(* IEC 61131-3 sources: kns-pump-station/tests/POUs/Model/FB_VfdSim_Test, 29 files *)

(* ---- FB_VfdSim_Test.decl.st ---- *)
// Назначение: набор coUnit для FB_VfdSim — модель ПЧ по условной карте: рампа к заданию и торможение, реле
//             «Работа», авария с выбегом и сброс по фронту CTW.2, коды аварий, потеря связи (регистры замирают,
//             записи не доходят), сторожевой таймер 5 с → 50 Гц (04 §12, PMI-28, PMI-29), восстановление связи,
//             пропадание питания и загрузка, инъекции ОС, местный пуск (частота местного поста), ток в регистре,
//             «время назад».
//             Время — PL.FB_FakeTime, шаг 100 мс; разгон 0 → 50 Гц за 10 с (5 Гц/с).
// Автор:      kr0nsch
// Версия:     0.1.0
// Документ:   docs/DESIGN.md, разделы 11.3, 14.1
FUNCTION_BLOCK FB_VfdSim_Test EXTENDS coUnit.FB_TestSuite
VAR CONSTANT
    T_STEP : TIME := T#100MS;
    UI_1S : UINT := 10;               // шагов в 1 с
    R_EPS_HZ : REAL := 1.0E-3;
    UI_FREF_50HZ : UINT := 5000;      // 0,01 Гц
    UI_FREF_30HZ : UINT := 3000;
    UI_FREF_25HZ : UINT := 2500;
    R_LOCAL_HZ : REAL := 50.0;        // частота местного поста (SIM_VFD_LOCAL_FREQ_HZ)
END_VAR

(* ---- CommLossFreezesRegisters.method.decl.st ---- *)
// Потеря связи на 25 Гц: xCommOk = FALSE, регистры STW и FACT замирают; новое задание не доходит
// (частота 25 Гц); стоп по проводу работает (через 2 с — 15 Гц), а FACT по-прежнему 2500.
METHOD PRIVATE CommLossFreezesRegisters
VAR
    fbTime : PL.FB_FakeTime;    // подменное время
    fbDut : FB_VfdSim;          // проверяемая модель ПЧ
    uiI : UINT;
END_VAR

(* ---- CommLossFreezesRegisters.method.impl.st ---- *)
coUnit.TEST('VfdSim_CommLossFreezesRegisters');

fbDut(xRunCmd := TRUE, uiFref := UI_FREF_25HZ, itfTime := fbTime);
FOR uiI := 1 TO 6 * UI_1S DO
    fbTime.Advance(tStep := T_STEP);
    fbDut(itfTime := fbTime);
END_FOR
AssertEquals_UINT(Expected := 2500, Actual := fbDut.uiFact, Message := 'FACT 2500 before loss');
fbDut.xCommLoss := TRUE;
FOR uiI := 1 TO 1 DO
    fbTime.Advance(tStep := T_STEP);
    fbDut(itfTime := fbTime);
END_FOR
AssertFalse(Condition := fbDut.xCommOk, Message := 'no comm');
fbDut.uiFref := UI_FREF_50HZ;
FOR uiI := 1 TO 2 * UI_1S DO
    fbTime.Advance(tStep := T_STEP);
    fbDut(itfTime := fbTime);
END_FOR
AssertEquals_REAL(Expected := 25.0, Actual := fbDut.rFreq_Hz, Delta := R_EPS_HZ,
                  Message := 'new reference not received');
fbDut.xRunCmd := FALSE;
FOR uiI := 1 TO 2 * UI_1S DO
    fbTime.Advance(tStep := T_STEP);
    fbDut(itfTime := fbTime);
END_FOR
AssertEquals_REAL(Expected := 15.0, Actual := fbDut.rFreq_Hz, Delta := R_EPS_HZ, Message := 'wired stop works');
AssertEquals_UINT(Expected := 2500, Actual := fbDut.uiFact, Message := 'FACT frozen');
AssertEquals_WORD(Expected := GVL_Const.VFD_STW_READY OR GVL_Const.VFD_STW_RUNNING OR GVL_Const.VFD_STW_REMOTE,
                  Actual := fbDut.wStw, Message := 'STW frozen');

coUnit.TEST_FINISHED();

(* ---- CommLossWatchdogGoesTo50HzAfter5s.method.decl.st ---- *)
// Сторожевой таймер ПЧ (04 §12): работающий на 30 Гц насос через 4,9 с без связи — ещё задание 30 Гц,
// в 5,0 с — 50 Гц, через 4 с разгона — 50 Гц. Стоящий насос без связи (последнее задание 0): пуск по
// проводу после срабатывания таймера — разгон до 50 Гц, а не работа на 0 Гц.
METHOD PRIVATE CommLossWatchdogGoesTo50HzAfter5s
VAR
    fbTime : PL.FB_FakeTime;    // подменное время
    fbDut : FB_VfdSim;          // проверяемая модель ПЧ
    uiI : UINT;
    fbStopped : FB_VfdSim;      // ПЧ стоящего насоса
END_VAR

(* ---- CommLossWatchdogGoesTo50HzAfter5s.method.impl.st ---- *)
coUnit.TEST('VfdSim_CommLossWatchdogGoesTo50HzAfter5s');

fbDut(xRunCmd := TRUE, uiFref := UI_FREF_30HZ, itfTime := fbTime);
fbStopped(xRunCmd := FALSE, uiFref := 0, itfTime := fbTime);
FOR uiI := 1 TO 6 * UI_1S DO
    fbTime.Advance(tStep := T_STEP);
    fbDut(itfTime := fbTime);
END_FOR
fbDut.xCommLoss := TRUE;
fbStopped.xCommLoss := TRUE;
fbTime.Advance(tStep := T_STEP);
fbDut(itfTime := fbTime);
fbStopped(itfTime := fbTime);
FOR uiI := 1 TO 5 * UI_1S - 1 DO
    fbTime.Advance(tStep := T_STEP);
    fbDut(itfTime := fbTime);
    fbStopped(itfTime := fbTime);
END_FOR
AssertFalse(Condition := fbDut.xWatchdog, Message := 'no watchdog at 4.9 s');
AssertEquals_REAL(Expected := 30.0, Actual := fbDut.rRef_Hz, Delta := R_EPS_HZ, Message := 'last reference 30 Hz');
fbTime.Advance(tStep := T_STEP);
fbDut(itfTime := fbTime);
fbStopped(itfTime := fbTime);
AssertTrue(Condition := fbDut.xWatchdog AND fbStopped.xWatchdog, Message := 'watchdog at 5.0 s');
AssertEquals_REAL(Expected := GVL_Const.SIM_VFD_WATCHDOG_FREQ_HZ, Actual := fbDut.rRef_Hz, Delta := 0.0,
                  Message := 'preset 50 Hz');
FOR uiI := 1 TO 10 * UI_1S DO
    fbTime.Advance(tStep := T_STEP);
    fbDut(itfTime := fbTime);
    fbStopped(xRunCmd := TRUE, itfTime := fbTime);
END_FOR
AssertEquals_REAL(Expected := 50.0, Actual := fbDut.rFreq_Hz, Delta := R_EPS_HZ, Message := 'running pump at 50 Hz');
AssertEquals_REAL(Expected := 50.0, Actual := fbStopped.rFreq_Hz, Delta := R_EPS_HZ,
                  Message := 'pump started by wire runs at 50 Hz');

coUnit.TEST_FINISHED();

(* ---- CommRestoredFollowsFref.method.decl.st ---- *)
// После срабатывания таймера (50 Гц) связь восстановлена с заданием 3000: таймер снят, задание 30 Гц,
// через 4 с — 30 Гц, регистры снова обновляются (FACT 3000).
METHOD PRIVATE CommRestoredFollowsFref
VAR
    fbTime : PL.FB_FakeTime;    // подменное время
    fbDut : FB_VfdSim;          // проверяемая модель ПЧ
    uiI : UINT;
END_VAR

(* ---- CommRestoredFollowsFref.method.impl.st ---- *)
coUnit.TEST('VfdSim_CommRestoredFollowsFref');

fbDut(xRunCmd := TRUE, uiFref := UI_FREF_50HZ, itfTime := fbTime);
FOR uiI := 1 TO 10 * UI_1S DO
    fbTime.Advance(tStep := T_STEP);
    fbDut(itfTime := fbTime);
END_FOR
fbDut.xCommLoss := TRUE;
FOR uiI := 1 TO 6 * UI_1S DO
    fbTime.Advance(tStep := T_STEP);
    fbDut(itfTime := fbTime);
END_FOR
AssertTrue(Condition := fbDut.xWatchdog, Message := 'watchdog active');
fbDut.xCommLoss := FALSE;
fbDut.uiFref := UI_FREF_30HZ;
FOR uiI := 1 TO 1 DO
    fbTime.Advance(tStep := T_STEP);
    fbDut(itfTime := fbTime);
END_FOR
AssertTrue(Condition := fbDut.xCommOk AND NOT fbDut.xWatchdog, Message := 'comm restored, watchdog off');
AssertEquals_REAL(Expected := 30.0, Actual := fbDut.rRef_Hz, Delta := R_EPS_HZ, Message := 'follows FREF again');
FOR uiI := 1 TO 4 * UI_1S DO
    fbTime.Advance(tStep := T_STEP);
    fbDut(itfTime := fbTime);
END_FOR
AssertEquals_REAL(Expected := 30.0, Actual := fbDut.rFreq_Hz, Delta := R_EPS_HZ, Message := 'ramped to 30 Hz');
AssertEquals_UINT(Expected := 3000, Actual := fbDut.uiFact, Message := 'FACT updated');

coUnit.TEST_FINISHED();

(* ---- CurrentRegisterScaled.method.decl.st ---- *)
// Ток двигателя в регистре 102 — 0,1 А: 26,38 А → 264; неконечный ток и стоящий ПЧ — 0.
METHOD PRIVATE CurrentRegisterScaled
VAR
    fbTime : PL.FB_FakeTime;    // подменное время
    fbDut : FB_VfdSim;          // проверяемая модель ПЧ
    uiI : UINT;
    uBits : PL.U_RealBits;
END_VAR

(* ---- CurrentRegisterScaled.method.impl.st ---- *)
coUnit.TEST('VfdSim_CurrentRegisterScaled');

fbDut(xRunCmd := TRUE, uiFref := UI_FREF_50HZ, itfTime := fbTime);
FOR uiI := 1 TO 10 * UI_1S DO
    fbTime.Advance(tStep := T_STEP);
    fbDut(itfTime := fbTime);
END_FOR
fbDut.rMotorCurrent_A := 26.38;
FOR uiI := 1 TO 1 DO
    fbTime.Advance(tStep := T_STEP);
    fbDut(itfTime := fbTime);
END_FOR
AssertEquals_UINT(Expected := 264, Actual := fbDut.uiCurrent, Message := '26.38 A -> 264');
uBits.dwValue := 16#7FC00000;
fbDut.rMotorCurrent_A := uBits.rValue;
FOR uiI := 1 TO 1 DO
    fbTime.Advance(tStep := T_STEP);
    fbDut(itfTime := fbTime);
END_FOR
AssertEquals_UINT(Expected := 0, Actual := fbDut.uiCurrent, Message := 'NaN current -> 0');
fbDut.rMotorCurrent_A := 26.38;
fbDut.xRunCmd := FALSE;
FOR uiI := 1 TO 11 * UI_1S DO
    fbTime.Advance(tStep := T_STEP);
    fbDut(itfTime := fbTime);
END_FOR
AssertEquals_UINT(Expected := 0, Actual := fbDut.uiCurrent, Message := 'stopped drive -> 0');

coUnit.TEST_FINISHED();

(* ---- DefaultsReadyAndStopped.method.decl.st ---- *)
// Первый вызов с питанием: ПЧ готов, связь есть, STW = готов + дистанционное (16#0011), частота и
// FACT 0, код аварии 0, реле разомкнуты.
METHOD PRIVATE DefaultsReadyAndStopped
VAR
    fbTime : PL.FB_FakeTime;    // подменное время
    fbDut : FB_VfdSim;          // проверяемая модель ПЧ
END_VAR

(* ---- FaultCoastAndResetEdge.method.decl.st ---- *)
// Авария ПЧ на 50 Гц: выбег (частота 0 сразу), реле «Авария», STW.2, код 11, не готов. Сброс при
// активной инъекции не снимает; после снятия инъекции нужен новый фронт CTW.2; код аварии остаётся.
METHOD PRIVATE FaultCoastAndResetEdge
VAR
    fbTime : PL.FB_FakeTime;    // подменное время
    fbDut : FB_VfdSim;          // проверяемая модель ПЧ
    uiI : UINT;
END_VAR

(* ---- FaultCoastAndResetEdge.method.impl.st ---- *)
coUnit.TEST('VfdSim_FaultCoastAndResetEdge');

fbDut(xRunCmd := TRUE, uiFref := UI_FREF_50HZ, itfTime := fbTime);
FOR uiI := 1 TO 10 * UI_1S DO
    fbTime.Advance(tStep := T_STEP);
    fbDut(itfTime := fbTime);
END_FOR
fbDut.xFaultInj := TRUE;
FOR uiI := 1 TO 1 DO
    fbTime.Advance(tStep := T_STEP);
    fbDut(itfTime := fbTime);
END_FOR
AssertEquals_REAL(Expected := 0.0, Actual := fbDut.rFreq_Hz, Delta := 0.0, Message := 'coast: frequency 0');
AssertTrue(Condition := fbDut.xRelayFault AND fbDut.xFaulted AND NOT fbDut.xReady, Message := 'fault latched');
AssertFalse(Condition := fbDut.xRelayRun, Message := 'run relay open');
AssertEquals_WORD(Expected := GVL_Const.VFD_STW_FAULT OR GVL_Const.VFD_STW_REMOTE, Actual := fbDut.wStw,
                  Message := 'STW fault + remote');
AssertEquals_UINT(Expected := GVL_Const.SIM_VFD_FCODE_EXT, Actual := fbDut.uiFcode, Message := 'fault code 11');
fbDut.wCtw := GVL_Const.VFD_CTW_RESET;
FOR uiI := 1 TO 1 DO
    fbTime.Advance(tStep := T_STEP);
    fbDut(itfTime := fbTime);
END_FOR
AssertTrue(Condition := fbDut.xFaulted, Message := 'reset ignored while cause active');
fbDut.xFaultInj := FALSE;
FOR uiI := 1 TO 1 DO
    fbTime.Advance(tStep := T_STEP);
    fbDut(itfTime := fbTime);
END_FOR
AssertTrue(Condition := fbDut.xFaulted, Message := 'no new reset edge: still faulted');
fbDut.wCtw := 0;
FOR uiI := 1 TO 1 DO
    fbTime.Advance(tStep := T_STEP);
    fbDut(itfTime := fbTime);
END_FOR
fbDut.wCtw := GVL_Const.VFD_CTW_RESET;
FOR uiI := 1 TO 1 DO
    fbTime.Advance(tStep := T_STEP);
    fbDut(itfTime := fbTime);
END_FOR
AssertFalse(Condition := fbDut.xFaulted OR fbDut.xRelayFault, Message := 'reset edge clears fault');
AssertTrue(Condition := fbDut.xReady, Message := 'ready again');
AssertEquals_UINT(Expected := GVL_Const.SIM_VFD_FCODE_EXT, Actual := fbDut.uiFcode, Message := 'last fault code kept');
FOR uiI := 1 TO 1 DO
    fbTime.Advance(tStep := T_STEP);
    fbDut(itfTime := fbTime);
END_FOR
AssertTrue(Condition := fbDut.xOutputActive AND fbDut.rFreq_Hz > 0.0, Message := 'wired run restarts the drive');

coUnit.TEST_FINISHED();

(* ---- FeedbackStuckInjection.method.decl.st ---- *)
// Инъекция «ОС залипла»: ПЧ стоит, реле «Работа» замкнуто.
METHOD PRIVATE FeedbackStuckInjection
VAR
    fbTime : PL.FB_FakeTime;    // подменное время
    fbDut : FB_VfdSim;          // проверяемая модель ПЧ
END_VAR

(* ---- LocalRun.method.decl.st ---- *)
// «Местное»: провод «Пуск» от ПЛК не действует, пуск — с местного поста; бит STW.4 (дистанционное)
// снят.
METHOD PRIVATE LocalRun
VAR
    fbTime : PL.FB_FakeTime;    // подменное время
    fbDut : FB_VfdSim;          // проверяемая модель ПЧ
    uiI : UINT;
END_VAR

(* ---- LocalRun.method.impl.st ---- *)
coUnit.TEST('VfdSim_LocalRun');

fbDut(xRunCmd := TRUE, xLocal := TRUE, uiFref := UI_FREF_50HZ, itfTime := fbTime);
FOR uiI := 1 TO UI_1S DO
    fbTime.Advance(tStep := T_STEP);
    fbDut(itfTime := fbTime);
END_FOR
AssertFalse(Condition := fbDut.xOutputActive, Message := 'PLC wire ignored in local');
AssertEquals_WORD(Expected := GVL_Const.VFD_STW_READY, Actual := fbDut.wStw, Message := 'STW without remote bit');
fbDut.xLocalRun := TRUE;
FOR uiI := 1 TO UI_1S DO
    fbTime.Advance(tStep := T_STEP);
    fbDut(itfTime := fbTime);
END_FOR
AssertTrue(Condition := fbDut.xOutputActive AND fbDut.xRelayRun, Message := 'local run starts the drive');
AssertEquals_REAL(Expected := 5.0, Actual := fbDut.rFreq_Hz, Delta := R_EPS_HZ, Message := 'ramp in local');

coUnit.TEST_FINISHED();

(* ---- LocalRunAtLocalPreset.method.decl.st ---- *)
// «Местное», пуск по месту у стоящего насоса: FB_MotorVfd в Local держит задание равным фактической
// скорости (0 % у стоящего насоса), FREF = 0. ПЧ разгоняется к частоте местного поста (50 Гц) за tAccel,
// записи FREF мастера в «Местном» не действуют; после возврата в «Дистанционное» — снова FREF.
METHOD PRIVATE LocalRunAtLocalPreset
VAR
    fbTime : PL.FB_FakeTime;    // подменное время
    fbDut : FB_VfdSim;          // проверяемая модель ПЧ
    uiI : UINT;
END_VAR

(* ---- LocalRunAtLocalPreset.method.impl.st ---- *)
coUnit.TEST('VfdSim_LocalRunAtLocalPreset');

fbDut(xLocal := TRUE, xLocalRun := TRUE, uiFref := 0, itfTime := fbTime);
FOR uiI := 1 TO 10 * UI_1S DO
    fbTime.Advance(tStep := T_STEP);
    fbDut(itfTime := fbTime);
END_FOR
AssertTrue(Condition := fbDut.xOutputActive AND fbDut.xRelayRun, Message := 'local run starts the drive');
AssertEquals_REAL(Expected := R_LOCAL_HZ, Actual := fbDut.rFreq_Hz, Delta := R_EPS_HZ,
                  Message := 'local preset reached in tAccel');
fbDut.uiFref := UI_FREF_25HZ;
FOR uiI := 1 TO UI_1S DO
    fbTime.Advance(tStep := T_STEP);
    fbDut(itfTime := fbTime);
END_FOR
AssertEquals_REAL(Expected := R_LOCAL_HZ, Actual := fbDut.rFreq_Hz, Delta := R_EPS_HZ,
                  Message := 'master FREF ignored in local');
fbDut.xLocal := FALSE;
fbDut.xLocalRun := FALSE;
fbDut.xRunCmd := TRUE;
FOR uiI := 1 TO 5 * UI_1S DO
    fbTime.Advance(tStep := T_STEP);
    fbDut(itfTime := fbTime);
END_FOR
AssertEquals_REAL(Expected := 25.0, Actual := fbDut.rFreq_Hz, Delta := R_EPS_HZ, Message := 'remote: back to FREF');

coUnit.TEST_FINISHED();

(* ---- NoFeedbackInjection.method.decl.st ---- *)
// Инъекция «нет ОС»: ПЧ вращает насос, реле «Работа» разомкнуто.
METHOD PRIVATE NoFeedbackInjection
VAR
    fbTime : PL.FB_FakeTime;    // подменное время
    fbDut : FB_VfdSim;          // проверяемая модель ПЧ
    uiI : UINT;
END_VAR

(* ---- NoFeedbackInjection.method.impl.st ---- *)
coUnit.TEST('VfdSim_NoFeedbackInjection');

fbDut(xRunCmd := TRUE, uiFref := UI_FREF_50HZ, itfTime := fbTime);
FOR uiI := 1 TO 10 * UI_1S DO
    fbTime.Advance(tStep := T_STEP);
    fbDut(itfTime := fbTime);
END_FOR
fbDut.xNoFeedback := TRUE;
FOR uiI := 1 TO 1 DO
    fbTime.Advance(tStep := T_STEP);
    fbDut(itfTime := fbTime);
END_FOR
AssertTrue(Condition := fbDut.rFreq_Hz > 0.0 AND fbDut.xOutputActive, Message := 'drive running');
AssertFalse(Condition := fbDut.xRelayRun, Message := 'run relay open (no feedback)');

coUnit.TEST_FINISHED();

(* ---- OverheatFaultCode.method.decl.st ---- *)
// Перегрев (TS1n2 разрывает цепь аварии): авария ПЧ с кодом 12, выбег.
METHOD PRIVATE OverheatFaultCode
VAR
    fbTime : PL.FB_FakeTime;    // подменное время
    fbDut : FB_VfdSim;          // проверяемая модель ПЧ
    uiI : UINT;
END_VAR

(* ---- OverheatFaultCode.method.impl.st ---- *)
coUnit.TEST('VfdSim_OverheatFaultCode');

fbDut(xRunCmd := TRUE, uiFref := UI_FREF_50HZ, itfTime := fbTime);
FOR uiI := 1 TO 10 * UI_1S DO
    fbTime.Advance(tStep := T_STEP);
    fbDut(itfTime := fbTime);
END_FOR
fbDut.xOverheat := TRUE;
FOR uiI := 1 TO 1 DO
    fbTime.Advance(tStep := T_STEP);
    fbDut(itfTime := fbTime);
END_FOR
AssertTrue(Condition := fbDut.xFaulted AND fbDut.xRelayFault, Message := 'overheat trips the drive');
AssertEquals_UINT(Expected := GVL_Const.SIM_VFD_FCODE_OVERHEAT, Actual := fbDut.uiFcode, Message := 'fault code 12');
AssertEquals_REAL(Expected := 0.0, Actual := fbDut.rFreq_Hz, Delta := 0.0, Message := 'coast');

coUnit.TEST_FINISHED();

(* ---- PowerLossAndBoot.method.decl.st ---- *)
// Пропадание питания на ходу: частота 0, реле разомкнуты, связи нет, регистры 0. Питание вернулось
// (первый шаг цикла — вызов с питанием): 4,9 с ПЧ загружается (STW 0, связи нет), в 5,0 с готов, код
// последней аварии 13 (пониженное напряжение), пуск по проводу удержан — разгон.
METHOD PRIVATE PowerLossAndBoot
VAR
    fbTime : PL.FB_FakeTime;    // подменное время
    fbDut : FB_VfdSim;          // проверяемая модель ПЧ
    uiI : UINT;
END_VAR

(* ---- PowerLossAndBoot.method.impl.st ---- *)
coUnit.TEST('VfdSim_PowerLossAndBoot');

fbDut(xRunCmd := TRUE, uiFref := UI_FREF_50HZ, itfTime := fbTime);
FOR uiI := 1 TO 10 * UI_1S DO
    fbTime.Advance(tStep := T_STEP);
    fbDut(itfTime := fbTime);
END_FOR
fbDut.xPowerOk := FALSE;
FOR uiI := 1 TO 1 DO
    fbTime.Advance(tStep := T_STEP);
    fbDut(itfTime := fbTime);
END_FOR
AssertEquals_REAL(Expected := 0.0, Actual := fbDut.rFreq_Hz, Delta := 0.0, Message := 'no power: frequency 0');
AssertFalse(Condition := fbDut.xRelayRun OR fbDut.xCommOk OR fbDut.xReady, Message := 'no power: relays, comm off');
AssertEquals_WORD(Expected := 0, Actual := fbDut.wStw, Message := 'no power: STW 0');
fbDut.xPowerOk := TRUE;
FOR uiI := 1 TO 5 * UI_1S DO
    fbTime.Advance(tStep := T_STEP);
    fbDut(itfTime := fbTime);
END_FOR
AssertFalse(Condition := fbDut.xReady OR fbDut.xCommOk, Message := 'booting at 4.9 s');
AssertEquals_WORD(Expected := 0, Actual := fbDut.wStw, Message := 'booting: STW 0');
FOR uiI := 1 TO 1 DO
    fbTime.Advance(tStep := T_STEP);
    fbDut(itfTime := fbTime);
END_FOR
AssertTrue(Condition := fbDut.xReady AND fbDut.xCommOk, Message := 'ready after boot');
AssertEquals_UINT(Expected := GVL_Const.SIM_VFD_FCODE_UNDERVOLT, Actual := fbDut.uiFcode,
                  Message := 'last fault: undervoltage');
AssertTrue(Condition := fbDut.xOutputActive, Message := 'held wired run restarts after boot');

coUnit.TEST_FINISHED();

(* ---- RampToReference.method.decl.st ---- *)
// Пуск с заданием 5000 (50 Гц): через 5 с — 25 Гц (FACT 2500), через 10 с — 50 Гц; реле «Работа»
// и бит STW.1. Стоп: торможение 5 Гц/с, реле замкнуто до остановки (через 9,9 с — 0,5 Гц), в 10 с — 0.
METHOD PRIVATE RampToReference
VAR
    fbTime : PL.FB_FakeTime;    // подменное время
    fbDut : FB_VfdSim;          // проверяемая модель ПЧ
    uiI : UINT;
END_VAR

(* ---- RampToReference.method.impl.st ---- *)
coUnit.TEST('VfdSim_RampToReference');

fbDut(xRunCmd := TRUE, uiFref := UI_FREF_50HZ, itfTime := fbTime);
FOR uiI := 1 TO 5 * UI_1S DO
    fbTime.Advance(tStep := T_STEP);
    fbDut(itfTime := fbTime);
END_FOR
AssertEquals_REAL(Expected := 25.0, Actual := fbDut.rFreq_Hz, Delta := R_EPS_HZ, Message := '25 Hz after 5 s');
AssertEquals_UINT(Expected := 2500, Actual := fbDut.uiFact, Message := 'FACT 2500');
AssertTrue(Condition := fbDut.xRelayRun, Message := 'run relay closed');
AssertEquals_WORD(Expected := GVL_Const.VFD_STW_READY OR GVL_Const.VFD_STW_RUNNING OR GVL_Const.VFD_STW_REMOTE,
                  Actual := fbDut.wStw, Message := 'STW ready + running + remote');
FOR uiI := 1 TO 5 * UI_1S DO
    fbTime.Advance(tStep := T_STEP);
    fbDut(itfTime := fbTime);
END_FOR
AssertEquals_REAL(Expected := 50.0, Actual := fbDut.rFreq_Hz, Delta := R_EPS_HZ, Message := '50 Hz after 10 s');
AssertEquals_UINT(Expected := 5000, Actual := fbDut.uiFact, Message := 'FACT 5000');
fbDut.xRunCmd := FALSE;
FOR uiI := 1 TO 10 * UI_1S - 1 DO
    fbTime.Advance(tStep := T_STEP);
    fbDut(itfTime := fbTime);
END_FOR
AssertEquals_REAL(Expected := 0.5, Actual := fbDut.rFreq_Hz, Delta := R_EPS_HZ, Message := 'decelerating: 0.5 Hz');
AssertTrue(Condition := fbDut.xRelayRun, Message := 'run relay closed while decelerating');
FOR uiI := 1 TO 1 DO
    fbTime.Advance(tStep := T_STEP);
    fbDut(itfTime := fbTime);
END_FOR
AssertEquals_REAL(Expected := 0.0, Actual := fbDut.rFreq_Hz, Delta := 0.0, Message := 'stopped');
AssertFalse(Condition := fbDut.xRelayRun OR fbDut.xOutputActive, Message := 'run relay open after stop');

coUnit.TEST_FINISHED();

(* ---- ResetDriveClearsFault.method.decl.st ---- *)
// ResetDrive («ПЧ готовы», xResetPlant) снимает аварию, если причины уже нет, без фронта CTW.2;
// при активной причине авария остаётся.
METHOD PRIVATE ResetDriveClearsFault
VAR
    fbTime : PL.FB_FakeTime;    // подменное время
    fbDut : FB_VfdSim;          // проверяемая модель ПЧ
    uiI : UINT;
END_VAR

(* ---- ResetDriveClearsFault.method.impl.st ---- *)
coUnit.TEST('VfdSim_ResetDriveClearsFault');

fbDut(xRunCmd := TRUE, uiFref := UI_FREF_50HZ, itfTime := fbTime);
FOR uiI := 1 TO 10 * UI_1S DO
    fbTime.Advance(tStep := T_STEP);
    fbDut(itfTime := fbTime);
END_FOR
fbDut.xFaultInj := TRUE;
FOR uiI := 1 TO 1 DO
    fbTime.Advance(tStep := T_STEP);
    fbDut(itfTime := fbTime);
END_FOR
fbDut.ResetDrive();
FOR uiI := 1 TO 1 DO
    fbTime.Advance(tStep := T_STEP);
    fbDut(itfTime := fbTime);
END_FOR
AssertTrue(Condition := fbDut.xFaulted, Message := 'cause active: fault stays');
fbDut.xFaultInj := FALSE;
fbDut.ResetDrive();
FOR uiI := 1 TO 1 DO
    fbTime.Advance(tStep := T_STEP);
    fbDut(itfTime := fbTime);
END_FOR
AssertFalse(Condition := fbDut.xFaulted, Message := 'ResetDrive clears fault');
AssertTrue(Condition := fbDut.xReady, Message := 'ready');

coUnit.TEST_FINISHED();

(* ---- TimeBackwardsHoldsFrequency.method.decl.st ---- *)
// «Время назад»: шаг рампы 0 — частота не меняется; дальше рампа продолжается.
METHOD PRIVATE TimeBackwardsHoldsFrequency
VAR
    fbTime : PL.FB_FakeTime;    // подменное время
    fbDut : FB_VfdSim;          // проверяемая модель ПЧ
    uiI : UINT;
END_VAR

(* ---- TimeBackwardsHoldsFrequency.method.impl.st ---- *)
coUnit.TEST('VfdSim_TimeBackwardsHoldsFrequency');

fbDut(xRunCmd := TRUE, uiFref := UI_FREF_50HZ, itfTime := fbTime);
FOR uiI := 1 TO 3 * UI_1S DO
    fbTime.Advance(tStep := T_STEP);
    fbDut(itfTime := fbTime);
END_FOR
AssertEquals_REAL(Expected := 15.0, Actual := fbDut.rFreq_Hz, Delta := R_EPS_HZ, Message := '15 Hz after 3 s');
fbTime.SetNow(ltValue := fbTime.Now() - LTIME#1S);
fbDut(itfTime := fbTime);
AssertEquals_REAL(Expected := 15.0, Actual := fbDut.rFreq_Hz, Delta := R_EPS_HZ,
                  Message := 'time back: frequency held');
FOR uiI := 1 TO 1 DO
    fbTime.Advance(tStep := T_STEP);
    fbDut(itfTime := fbTime);
END_FOR
AssertEquals_REAL(Expected := 15.5, Actual := fbDut.rFreq_Hz, Delta := R_EPS_HZ, Message := 'ramp resumes');

coUnit.TEST_FINISHED();
